(* IEC 61131-3 sources: ironplc/compiler/plc2plc/resources/test, 32 files *)

(* ---- sized_string_contexts_rendered.st ---- *)
FUNCTION FUNC_WITH_VAR_STRING : INT
   VAR_INPUT
      x : INT;
   END_VAR

   VAR
      buf : STRING [ 10 ];
   END_VAR

   VAR
      wbuf : WSTRING [ 20 ];
   END_VAR

   FUNC_WITH_VAR_STRING := 0 ;
END_FUNCTION
FUNCTION FUNC_WITH_VAR_CONSTANT_STRING : INT
   VAR CONSTANT
      FILL : STRING [ 1 ] :='0';
   END_VAR

   VAR CONSTANT
      WFILL : WSTRING [ 1 ] :="0";
   END_VAR

   FUNC_WITH_VAR_CONSTANT_STRING := 0 ;
END_FUNCTION
FUNCTION FUNC_WITH_VAR_IN_OUT_STRING : INT
   VAR_IN_OUT
      buf : STRING [ 255 ];
   END_VAR

   VAR_IN_OUT
      wbuf : WSTRING [ 255 ];
   END_VAR

   FUNC_WITH_VAR_IN_OUT_STRING := 0 ;
END_FUNCTION
TYPE
   STRUCT_WITH_STRING : STRUCT
      name : STRING [ 10 ] ;
      wname : WSTRING [ 20 ] ;
   END_STRUCT ;
END_TYPE

(* ---- strings_rendered.st ---- *)
TYPE
   TEXT_EXTENDED : STRING [ 1 ] :='�' ;
END_TYPE

(* ---- type_decl_rendered.st ---- *)
TYPE
   VALUES_ENUM : ( VAL1 , VAL2 , VAL3 ) ;
END_TYPE
TYPE
   VALUES_ENUM_WITH_DEFAULT : ( VAL1 , VAL2 , VAL3 ) := VAL2 ;
END_TYPE
TYPE
   LIMIT_RANGE : UINT ( 0.. 3 ) ;
END_TYPE
TYPE
   LIMIT_RANGE_DEFAULT : UINT ( 0.. 3 ) := 1 ;
END_TYPE
TYPE
   LIMIT_RANGE_NEGATIVE : INT ( -10.. 10 ) ;
END_TYPE
TYPE
   ARR_RANGE : ARRAY [ 1.. 8 ] OF INT ;
END_TYPE
TYPE
   ARR_RANGE_2D : ARRAY [ 1.. 8 , 1.. 4 ] OF INT ;
END_TYPE
TYPE
   ARR_RANGE_ENUM : ARRAY [ 2.. 4 ] OF CUSTOM ;
END_TYPE
TYPE
   TEXT_EMPTY : STRING [ 1 ] ;
END_TYPE
TYPE
   TEXT_DEFAULT : STRING [ 5 ] :='value' ;
END_TYPE
TYPE
   WTEXT_EMPTY : WSTRING [ 1 ] ;
END_TYPE
TYPE
   WTEXT_DEFAULT : WSTRING [ 5 ] :="value" ;
END_TYPE
TYPE
   CUSTOM_STRUCT : STRUCT
      NAME : BOOL ;
   END_STRUCT ;
END_TYPE
TYPE
   CUSTOM_STRUCT_WITH_ENUM : STRUCT
      NAME : VAL_TYPE := INIT_VAL ;
      ARR_RANGE_ENUM : ARRAY [ 2.. 4 ] OF CUSTOM ;
      LIMIT_RANGE : UINT ( 0.. 3 ) ;
   END_STRUCT ;
END_TYPE
TYPE
   STR_WITH_SIZE : STRING [ 5 ] ;
END_TYPE
TYPE
   STR_WITH_SIZE_COMPATIBILITY : STRING [ 5 ] ;
END_TYPE

(* ---- array_in_function_var_rendered.st ---- *)
FUNCTION MY_FUNC : BOOL
   VAR_INPUT
      x : INT;
   END_VAR

   VAR
      stack : ARRAY [ 1.. 32 ] OF UINT;
   END_VAR

   stack[ 1 ] := INT_TO_UINT ( x ) ;
   MY_FUNC := BOOL#TRUE ;
END_FUNCTION

(* ---- array_of_string_rendered.st ---- *)
FUNCTION fun : BOOL
   VAR_INPUT
      names : ARRAY [ 1.. 3 ] OF STRING [ 10 ];
   END_VAR

   fun := BOOL#TRUE ;
END_FUNCTION

(* ---- array_rendered.st ---- *)
FUNCTION fun : BOOL
   VAR_INPUT
      var1 : INT;
   END_VAR

   VAR_INPUT
      pt : ARRAY [ 1.. 8 ] OF INT;
   END_VAR

   var1 := ( var1 + pt[ i ] ) ;
END_FUNCTION

(* ---- empty_var_block_rendered.st ---- *)
FUNCTION myFunc : INT
   VAR_INPUT
      x : INT;
   END_VAR

   myFunc := x ;
END_FUNCTION

(* ---- expressions_rendered.st ---- *)
FUNCTION fun : BOOL
   VAR_INPUT
      var1 : BYTE;
   END_VAR

   IF ( var1 < BYTE#32 ) THEN
      var1 := 1 ;
   END_IF ;

   var1 := NOT ( var3 OR var3 ) ;
   var1 := FUNC_NAME ( var1 , '  ' ) ;
   var1 := ( ( - 1 + ( 2 * 3 ) ) - ( ( 4 / 6 ) MOD ( 7 ** 8 ) ) ) ;
   var1 := ( ( ( ( 1 >= 2 ) <= 3 ) <> 4 ) XOR 5 ) ;
   IF ( var1 > TIME#1000ms ) THEN
      var1 := 1 ;
   END_IF ;

END_FUNCTION

(* ---- inout_var_decl_rendered.st ---- *)
FUNCTION FUNC : UINT
   VAR_IN_OUT
      E : REAL;
   END_VAR

   VAR_IN_OUT
      RNG : INT ( 1.. 2 );
   END_VAR

   VAR_IN_OUT
      ARR : ARRAY [ 0.. 3 ] OF INT;
   END_VAR

   array_avg := ( array_avg + arr[ idx ][ idx ] ) ;
END_FUNCTION

(* ---- input_var_decl_rendered.st ---- *)
FUNCTION FUNC : UINT
   VAR_INPUT
      E : REAL;
   END_VAR

   VAR_INPUT
      PI : BOOL R_EDGE;
   END_VAR

   VAR_INPUT
      G : BOOL R_EDGE;
   END_VAR

   array_avg := ( array_avg + arr[ idx ][ idx ] ) ;
END_FUNCTION

(* ---- nested_rendered.st ---- *)
FUNCTION fun : BOOL
   VAR_INPUT
      var1 : BYTE;
   END_VAR

   array_avg := ( array_avg + arr[ idx ][ idx ] ) ;
END_FUNCTION

(* ---- conditional_rendered.st ---- *)
FUNCTION_BLOCK BLOCK
   IF ( NOT VAR1 AND VAR1 ) THEN
      VAR1 := 1 ;
   ELSIF ( NOT VAR1 AND VAR1 ) THEN
      VAR1 := 1 ;
   END_IF ;

END_FUNCTION_BLOCK

(* ---- literal_rendered.st ---- *)
FUNCTION_BLOCK BLOCK

   VAR
      REAL_WITH_TYPE : REAL := LREAL#11.0;
   END_VAR

   VAR
      BOOL_WITH_TYPE_TRUE : BOOL := BOOL#TRUE;
   END_VAR

   VAR
      TOD_WITH_VALUE_INTEGRAL : TIME_OF_DAY := TIME_OF_DAY#14:30:20;
   END_VAR

   VAR
      DATE_WITH_VALUE : DATE := DATE#2024-01-20;
   END_VAR

   VAR
      DATE_AND_TIME_WITH_VALUE : DATE_AND_TIME := DATE_AND_TIME#2024-01-20-15:30:22;
   END_VAR
   REAL_WITH_TYPE := 10 ;

END_FUNCTION_BLOCK

(* ---- member_initializers.st ---- *)
TYPE
   Color : ( Red , Green ) ;
END_TYPE
TYPE
   Inner : STRUCT
      c : Color ;
   END_STRUCT ;
END_TYPE
TYPE
   Outer : STRUCT
      values : ARRAY [ 1.. 2 ] OF INT ;
      inner : Inner ;
   END_STRUCT ;
END_TYPE
FUNCTION_BLOCK Lamp

   VAR_INPUT
      color : Color;
   END_VAR

END_FUNCTION_BLOCK
PROGRAM main

VAR
   o : Outer := ( values := [ 1 , 2 ] , inner := ( c := Green ) );
END_VAR

VAR
   lamp : Lamp := ( color := Red );
END_VAR
END_PROGRAM

(* ---- oop_rendered.st ---- *)
INTERFACE I_Loggable
END_INTERFACE
INTERFACE I_Nameable
END_INTERFACE
INTERFACE I_Drivable EXTENDS I_Loggable
END_INTERFACE
FUNCTION_BLOCK ABSTRACT FB_BaseMotor IMPLEMENTS I_Drivable , I_Nameable

   VAR
      bRunning : BOOL;
   END_VAR

METHOD Start
   bRunning := BOOL#TRUE ;
END_METHOD
METHOD Stop
   bRunning := BOOL#FALSE ;
END_METHOD
END_FUNCTION_BLOCK
FUNCTION_BLOCK FB_ServoMotor EXTENDS FB_BaseMotor IMPLEMENTS I_Drivable

   VAR
      rSpeed : REAL;
   END_VAR

   VAR
      aHistory : ARRAY [ 0.. 3 ] OF REAL;
   END_VAR

METHOD SetSpeed : BOOL

   VAR_INPUT
      rNewSpeed : REAL;
   END_VAR

   SUPER^. Start ( ) ;
   rSpeed := rNewSpeed ;
   THIS^.aHistory[ 0 ] := rNewSpeed ;
   SetSpeed := BOOL#TRUE ;
END_METHOD
METHOD LogState
   IF SUPER^.bRunning THEN
      aHistory[ 1 ] := rSpeed ;
   END_IF ;

END_METHOD
METHOD Reset
   THIS^.rSpeed := 0.0 ;
   THIS^. LogState ( ) ;
   SUPER^. Stop ( ) ;
END_METHOD
END_FUNCTION_BLOCK
PROGRAM main

VAR
   m : FB_ServoMotor;
END_VAR
m. SetSpeed ( 1.5 ) ;
m. SetSpeed ( rNewSpeed := 2.0 ) ;
m. Reset ( ) ;
END_PROGRAM

(* ---- partial_access_bit_rendered.st ---- *)
FUNCTION_BLOCK MyBlock

   VAR
      myWord : WORD;
   END_VAR

   VAR
      myBool : BOOL;
   END_VAR
   myBool := myWord.0 ;
   myBool := myWord.15 ;

END_FUNCTION_BLOCK

(* ---- sfc_rendered.st ---- *)
FUNCTION_BLOCK sfc

   VAR_INPUT
      IN : BOOL;
   END_VAR

   VAR_OUTPUT
      OUT : INT;
   END_VAR

   VAR
      COUNT : INT;
   END_VAR
   INITIAL_STEP Start :
      RESET ( N );
   END_STEP

   TRANSITION FROM Start TO MidStep
      := BOOL#FALSE ;
   END_TRANSITION

   STEP MidStep :
      RESET ( N );
   END_STEP

   ACTION RESET :
      COUNT := 0 ;
   END_ACTION

END_FUNCTION_BLOCK

(* ---- textual_rendered.st ---- *)
FUNCTION_BLOCK BLOCK
   NUM_INT := 10 ;
   NUM_FLOAT := 10.0 ;
   IF ( NUM1 < NUM2 ) THEN
      NUM1 := 1 ;
   ELSIF ( NUM2 = NUM3 ) THEN
      NUM1 := 2 ;
   ELSE
      NUM1 := 3 ;
   END_IF ;

   CASE EXPR_WITH_ELSE OF
      VAL1 :
         (* empty *) ;
      VAL2 :
         NUM1 := 1 ;
      ELSE
         NUM2 := 2 ;
   END_CASE ;

   CASE EXPR_NO_ELSE OF
      VAL1 :
         (* empty *) ;
      VAL2 :
         NUM1 := 1 ;
   END_CASE ;

   FOR VAL1 := 1 TO 10 BY 1 DO
      VAL2 := VAL1 ;
   END_FOR ;

   WHILE ( VAL1 = 1 ) DO
      VAL2 := VAL1 ;
   END_WHILE ;

   REPEAT
      VAL2 := VAL1 ;
   UNTIL ( VAL2 = 2 )
   END_REPEAT ;

END_FUNCTION_BLOCK

(* ---- var_temp_rendered.st ---- *)
FUNCTION my_func : DINT
   VAR_INPUT
      a : DINT;
   END_VAR

   VAR_TEMP
      temp : DINT;
   END_VAR

   temp := ( a * 2 ) ;
   my_func := temp ;
END_FUNCTION
FUNCTION_BLOCK my_fb

   VAR_TEMP
      t : INT;
   END_VAR
   t := 42 ;

END_FUNCTION_BLOCK
PROGRAM main

VAR
   q : INT;
END_VAR

VAR_TEMP
   t : INT := 3;
END_VAR
q := t ;
END_PROGRAM

(* ---- adr_rendered.st ---- *)
PROGRAM main

VAR
   counter : INT := 42;
END_VAR

VAR
   p : POINTER TO INT;
END_VAR

VAR
   value : INT;
END_VAR
p := ADR ( counter ) ;
value := p^ ;
p^ := 99 ;
END_PROGRAM

(* ---- configuration_rendered.st ---- *)
CONFIGURATION config
   RESOURCE resource1 ON PLC
      TASK plc_task ( INTERVAL := TIME#100ms , PRIORITY := 1 ) ;
      PROGRAM plc_task_instance WITH plc_task : plc_prg ;
   END_RESOURCE
   VAR_CONFIG
Some.FunctionBlock.Item.Path : FB_TYPE_NAME := ( ELEM := VAL ) ;
Some.Located.Item.Path AT %QB1 : BYTE ;
   END_VAR

END_CONFIGURATION
PROGRAM main

VAR
   Button AT %IX1 : BOOL;
END_VAR

VAR
   Buzzer AT %QX1 : BOOL;
END_VAR
Buzzer := NOT Button ;
END_PROGRAM

(* ---- expression_types.st ---- *)
TYPE
    Color : (Red, Green, Blue);
END_TYPE

FUNCTION Scale : LREAL
VAR_INPUT
    raw : DINT;
    gain : LREAL;
END_VAR
    Scale := raw * gain;
END_FUNCTION

PROGRAM main
VAR
    count : INT;
    total : DINT;
    big : LINT;
    level : REAL;
    out : LREAL;
    flag : BOOL;
    arr : ARRAY[1..4] OF INT;
    i : INT;
    c : Color;
    elapsed : TIME;
    name : STRING[20];
    r : REF_TO INT;
END_VAR
    count := count + 1;
    flag := big > total;
    level := count;
    out := Scale(raw := total, gain := 0.5);
    FOR i := 1 TO 4 DO
        arr[i] := MAX(arr[i], count);
    END_FOR;
    IF NOT flag AND total < 10 THEN
        big := ABS(big) + total;
    END_IF;
    c := Green;
    flag := c = Red;
    elapsed := elapsed + T#1s;
    name := CONCAT(name, 'abc');
    r := REF(count);
    count := r^ + 1;
    r := NULL;
    count := INT#5 + 7;
END_PROGRAM

(* ---- expression_types_rendered.st ---- *)
TYPE
   Color : ( Red , Green , Blue ) ;
END_TYPE
FUNCTION Scale : LREAL
   VAR_INPUT
      raw : dint;
   END_VAR

   VAR_INPUT
      gain : lreal;
   END_VAR

   Scale := ( raw (* DINT -> LREAL *) * gain (* LREAL *) ) (* LREAL *) ;
END_FUNCTION
PROGRAM main

VAR
   count : int;
END_VAR

VAR
   total : dint;
END_VAR

VAR
   big : lint;
END_VAR

VAR
   level : real;
END_VAR

VAR
   out : lreal;
END_VAR

VAR
   flag : bool;
END_VAR

VAR
   arr : ARRAY [ 1.. 4 ] OF INT;
END_VAR

VAR
   i : int;
END_VAR

VAR
   c : Color;
END_VAR

VAR
   elapsed : time;
END_VAR

VAR
   name : STRING [ 20 ];
END_VAR

VAR
   r : REF_TO INT;
END_VAR
count := ( count (* INT *) + 1 (* CONSTANT INT *) ) (* INT *) ;
flag := ( big (* LINT *) > total (* DINT -> LINT *) ) (* BOOL *) ;
level := count (* INT -> REAL *) ;
out := Scale ( raw := total (* DINT *) , gain := 0.5 (* CONSTANT LREAL *) ) (* LREAL *) ;
FOR i := 1 (* CONSTANT INT *) TO 4 (* CONSTANT INT *) DO
   arr[ i (* INT *) ] := MAX ( IN1 := arr[ i (* INT *) ] (* INT *) , IN2 := count (* INT *) ) (* INT *) ;
END_FOR ;

IF ( ( NOT flag (* BOOL *) ) (* BOOL *) AND ( total (* DINT *) < 10 (* CONSTANT DINT *) ) (* BOOL *) ) (* BOOL *) THEN
   big := ( ABS ( IN := big (* LINT *) ) (* LINT *) + total (* DINT -> LINT *) ) (* LINT *) ;
END_IF ;

c := Green (* CONSTANT Color *) ;
flag := ( c (* Color *) = Red (* CONSTANT Color *) ) (* BOOL *) ;
elapsed := ( elapsed (* TIME *) + TIME#1000ms (* CONSTANT TIME *) ) (* TIME *) ;
name := CONCAT ( IN1 := name (* STRING *) , IN2 := 'abc' (* CONSTANT STRING *) ) (* STRING *) ;
r := REF( count ) (* REF_TO INT *) ;
count := ( ( r (* REF_TO INT *)^ ) (* INT *) + 1 (* CONSTANT INT *) ) (* INT *) ;
r := NULL (* CONSTANT NULL *) ;
count := 12 (* CONSTANT INT *) ;
END_PROGRAM

(* ---- partial_access_multi_rendered.st ---- *)
PROGRAM main

VAR
   d : DWORD;
END_VAR

VAR
   l : LWORD;
END_VAR

VAR
   rb : BYTE;
END_VAR

VAR
   rw : WORD;
END_VAR

VAR
   rd : DWORD;
END_VAR
rb := d.%B0 ;
rw := d.%W1 ;
rd := l.%D0 ;
d.%B2 := BYTE#255 ;
l.%W3 := WORD#43981 ;
END_PROGRAM

(* ---- pointer_to_rendered.st ---- *)
TYPE
   IntPtr : POINTER TO INT ;
END_TYPE
PROGRAM main

VAR
   counter : INT := 42;
END_VAR

VAR
   p : POINTER TO INT;
END_VAR

VAR
   ptrs : ARRAY [ 0.. 2 ] OF POINTER TO INT;
END_VAR

VAR
   value : INT;
END_VAR
p := REF( counter ) ;
value := p^ ;
p^ := 99 ;
p := NULL ;
END_PROGRAM

(* ---- program_rendered.st ---- *)
PROGRAM main

VAR
   Button AT %IX1 : BOOL;
END_VAR

VAR
   Buzzer AT %QX1 : BOOL;
END_VAR

VAR_ACCESS
   VarPath : VarName.Path : BOOL READ_ONLY;
END_VAR
Buzzer := NOT Button ;
END_PROGRAM

(* ---- ref_rendered.st ---- *)
TYPE
   IntRef : REF_TO INT ;
END_TYPE
TYPE
   ArrRef : REF_TO ARRAY [ 0.. 3 ] OF DINT ;
END_TYPE
FUNCTION read_ref : INT
   VAR_INPUT
      pt : REF_TO INT;
   END_VAR

   read_ref := pt^ ;
END_FUNCTION
PROGRAM main

VAR
   counter : INT := 42;
END_VAR

VAR
   r : REF_TO INT := REF( counter );
END_VAR

VAR
   r_null : REF_TO INT := NULL;
END_VAR

VAR
   r_uninit : REF_TO INT;
END_VAR

VAR
   data : REF_TO ARRAY [ 0.. 3 ] OF INT;
END_VAR

VAR
   refs : ARRAY [ 0.. 2 ] OF REF_TO INT;
END_VAR

VAR
   value : INT;
END_VAR
value := r^ ;
r^ := 99 ;
r := REF( counter ) ;
IF ( r <> NULL ) THEN
   value := r^ ;
END_IF ;

value := read_ref ( pt := REF( counter ) ) ;
END_PROGRAM

(* ---- reference_to_rendered.st ---- *)
TYPE
   IntRef : REFERENCE TO INT ;
END_TYPE
PROGRAM main

VAR
   counter : INT := 42;
END_VAR

VAR
   r : REFERENCE TO INT;
END_VAR

VAR
   refs : ARRAY [ 0.. 2 ] OF REFERENCE TO INT;
END_VAR

VAR
   value : INT;
END_VAR
r REF= counter ;
value := r^ ;
r^ := 99 ;
refs[ 0 ] REF= counter ;
value := refs[ 0 ]^ ;
END_PROGRAM

(* ---- sizeof_rendered.st ---- *)
PROGRAM main

VAR
   x : INT;
END_VAR

VAR
   y : DWORD;
END_VAR

VAR
   arr : ARRAY [ 1.. 10 ] OF INT;
END_VAR

VAR
   s : DINT;
END_VAR
s := SIZEOF ( x ) ;
s := SIZEOF ( y ) ;
s := SIZEOF ( arr ) ;
END_PROGRAM

(* ---- time_function_decl_rendered.st ---- *)
FUNCTION TIME : TIME TIME := TIME#0ms ;
END_FUNCTION
PROGRAM main

VAR
   t : TIME;
END_VAR
t := TIME ( ) ;
END_PROGRAM

(* ---- var_decl_rendered.st ---- *)
PROGRAM fb

VAR CONSTANT
   E : REAL := 2.718;
END_VAR

VAR
   AT %IX1.1 : BOOL;
END_VAR

VAR
   AT %IX2.1 : BOOL := 1;
END_VAR

VAR
   AT %MW1 : INT := 2;
END_VAR

VAR RETAIN
   AT %QW1 : WORD := 65280;
END_VAR

VAR RETAIN
   AT %QB2 : WORD := 4032;
END_VAR

VAR RETAIN
   AT %QB3 : WORD := 10;
END_VAR

VAR RETAIN
   C3 AT %MW1.2.3 : WORD;
END_VAR

VAR RETAIN
   C2 AT %Q* : BYTE;
END_VAR

VAR
   XWORD : INT;
END_VAR

VAR
   YWORD : INT;
END_VAR

VAR
   ZWORD : INT;
END_VAR

VAR
   UNINIT : ARRAY [ 0.. 9 ] OF INT;
END_VAR

VAR
   INIT : ARRAY [ 1.. 12 ] OF SINT := [ 2 , 7 , 18 ];
END_VAR

VAR
   MULTI_DIM_ARRAY : ARRAY [ 1.. 2 , 3.. 4 , 5.. 6 ] OF SINT;
END_VAR

VAR
   PARENTHESIS_ARRAY : ARRAY [ 0.. 3 ] OF SINT := [ 3 ( 2 ) ];
END_VAR

VAR
   VAL_STR : STRING [ 2 ];
END_VAR

VAR
   VAL_STR_INIT : STRING :='abc';
END_VAR

VAR
   VAL_STR_PREFIX : STRING :='ABC';
END_VAR

VAR
   VAL_STR_SIZED_INIT : STRING [ 3 ] :='abc';
END_VAR

VAR
   VAL_WSTR : WSTRING [ 9 ];
END_VAR

VAR
   VAL_WSTR_INIT : WSTRING :="def";
END_VAR

VAR
   VAL_WSTR_PREFIX : WSTRING :="ABC";
END_VAR

VAR
   VAL_WSTR_SIZED_INIT : WSTRING [ 3 ] :="def";
END_VAR

VAR
   NAME : ONE_STRUCT_ELEMENT := ( ELEM := VAL );
END_VAR

VAR
   NAME2 : TWO_STRUCT_ELEMENTS := ( ELEM1 := VAL1 , ELEM2 := VAL2 );
END_VAR

VAR
   NAME3 : STRUCT_TWO_ELEMENTS := ( ELEM1 := VAL1 , ELEM2 := VAL2 );
END_VAR

VAR
   X : REAL2;
END_VAR

VAR
   Y : REAL;
END_VAR
END_PROGRAM

(* ---- wstring_ops_rendered.st ---- *)
PROGRAM main

VAR
   a : WSTRING [ 10 ] :="foo";
END_VAR

VAR
   b : WSTRING [ 10 ] :="bar";
END_VAR

VAR
   c : WSTRING [ 20 ];
END_VAR

VAR
   s : STRING [ 20 ];
END_VAR

VAR
   n : DINT;
END_VAR

VAR
   eq : BOOL;
END_VAR
c := a ;
c := "baz" ;
s := 'baz' ;
c := CONCAT ( a , b ) ;
n := LEN ( a ) ;
eq := ( a = b ) ;
END_PROGRAM
